FUNCTION_BLOCK FB_stringBuilder
VAR_INPUT
END_VAR
VAR
	bBuffer				:	ARRAY[0..PARAMETERS.uiMaxCharacters - 1] OF BYTE;
	bBufferOld			:	ARRAY[0..PARAMETERS.uiMaxCharacters - 1] OF BYTE;
	udiIndex			:	UDINT;
	udiIndexOld			:	UDINT;
	pbBuffer			:	POINTER TO BYTE		:=	ADR(bBuffer);
	pbBufferOld			:	POINTER TO BYTE		:=	ADR(bBufferOld);
END_VAR

METHOD AddChar : BOOL
VAR_INPUT
	byChar	:	BYTE;
END_VAR
IF CheckLength() THEN
	bBuffer[udiIndex]	:=	byChar;
	AddChar			:=	TRUE;
	IncrementIndex();
END_IF
END_METHOD

ACTION AddCloseBracket:
AddChar(41);
END_ACTION

ACTION AddColon:
AddChar(58);
END_ACTION

ACTION AddComma:
AddChar(44);
END_ACTION

ACTION AddDollar:
AddChar(36);
END_ACTION

ACTION AddDot:
AddChar(46);
END_ACTION

ACTION AddDoubleQuote:
AddChar(34);
END_ACTION

METHOD AddKeyValue : BOOL
VAR_INPUT
	psKey	:	POINTER TO STRING;
	psValue	:	POINTER TO STRING;
END_VAR
AddString(psKey);
AddColon();
AddString(psValue);
AddComma();
END_METHOD

ACTION AddNewLine:
AddChar(10);
END_ACTION

ACTION AddNullChar:
IF NOT CheckLength() THEN
	udiIndex	:=	PARAMETERS.uiMaxCharacters - 1;
END_IF
AddChar(0);
END_ACTION

ACTION AddOpenBracket:
AddChar(40);
END_ACTION

ACTION AddQuote:
AddChar(39);
END_ACTION

ACTION AddSemicolon:
AddChar(59);
END_ACTION

ACTION AddSpace:
AddChar(32);
END_ACTION

METHOD AddString : BOOL
VAR_INPUT
	psString		:	POINTER TO STRING;
END_VAR
VAR
	udiLen	:	UDINT;
END_VAR
udiLen	:=	(LEN2(psString));
IF CheckFinalLength(udiLen) THEN
	MEMCPY(pbBuffer + udiIndex, psString, udiLen);
	IncrementIndexVariable(udiLen);
	AddString	:=	TRUE;
END_IF
END_METHOD

ACTION AddTab:
AddChar(9);
END_ACTION

ACTION AddUnderscore:
AddChar(95);
END_ACTION

METHOD BuildString : BOOL
VAR_INPUT
	psString	:	POINTER TO STRING;
END_VAR
AddNullChar();
MEMCPY( psString, ADR(bBuffer), udiIndex );
END_METHOD

METHOD CheckFinalLength : BOOL
VAR_INPUT
	udiLen	:	UDINT;
END_VAR
CheckFinalLength	:=	(udiIndex + udiLen) < PARAMETERS.uiMaxCharacters;
END_METHOD

METHOD CheckLength : BOOL
VAR_INPUT
END_VAR
CheckLength	:=	CheckFinalLength(0);
END_METHOD

METHOD CheckMinimumLength : BOOL
VAR_INPUT
END_VAR
CheckMinimumLength	:=	udiIndex > 0;
END_METHOD

ACTION DecrementIndex:
IF CheckMinimumLength() THEN
	udiIndex	:=	udiIndex - 1;
END_IF
END_ACTION

METHOD DeleteChars : BOOL
VAR_INPUT
	udiNumChars	:	UDINT;
END_VAR
udiNumChars	:=	MIN(udiNumChars, udiIndex);
MEMSET(pbBuffer + (udiIndex - udiNumChars), 0, udiNumChars);
udiIndex := udiIndex - udiNumChars;
END_METHOD

ACTION IncrementIndex:
IncrementIndexVariable(1);
END_ACTION

METHOD IncrementIndexVariable : BOOL
VAR_INPUT
	udiIncrement	:	UDINT;
END_VAR
udiIndex	:=	udiIndex + udiIncrement;
END_METHOD

ACTION ResetBuffer:
IF CheckMinimumLength() THEN
	udiIndexOld	:=	udiIndex - 1;
	MEMSET(	ADR(bBufferOld), 0, PARAMETERS.uiMaxCharacters);
	MEMCPY( ADR(bBufferOld), ADR(bBuffer), udiIndexOld);
	
	ResetIndex();
	MEMSET(	ADR(bBuffer), 0, PARAMETERS.uiMaxCharacters);
END_IF
END_ACTION

ACTION ResetIndex:
udiIndex	:=	0;
END_ACTION

END_FUNCTION_BLOCK

(* stored: Version 1.1.0.1, ProductVersion 3.1.4024.9
   POU FB_stringBuilder: Id {26bce644-87e4-4374-b58f-9389bc582a26}, SpecialFunc None
   Folder ACTIONs: Id {99776992-d8a0-4ed4-aa61-350cfed19f86}
   Folder METHODs: Id {9a2113b2-3380-4328-be6b-be03ed0cc5a6}
   Method AddChar: Id {acb1b8e0-0207-4f46-8378-b68a295cf363}
   Action AddCloseBracket: Id {444bcdd4-ba94-4df4-ab4d-d2ec81607a8f}
   Action AddColon: Id {955d0969-09fd-4ef7-a5fc-925f1bf3fba6}
   Action AddComma: Id {f598045d-14ce-4e49-8860-6889173f446b}
   Action AddDollar: Id {62dc17c3-04a8-45e3-b384-0493539ef6bb}
   Action AddDot: Id {e44675ea-41f7-4475-a1a8-be67ad3f2ca2}
   Action AddDoubleQuote: Id {634a5359-7116-406e-b4c1-826d6bf2f6c9}
   Method AddKeyValue: Id {ea0220f5-ed5d-41e8-9b72-147e94feed33}
   Action AddNewLine: Id {c2c363a3-f640-4a66-9c2e-ae6cfdf7030a}
   Action AddNullChar: Id {41965dbb-6995-4e5e-9350-33895695746a}
   Action AddOpenBracket: Id {2ec56027-8c0a-434b-a7a8-c83c4f1f8e42}
   Action AddQuote: Id {a0d24b89-7c31-4ef3-9361-6e66114a55e2}
   Action AddSemicolon: Id {6e821915-2f2b-48e5-a2be-50c5a41a7f62}
   Action AddSpace: Id {efb50eb6-39f2-45ad-afb8-a2137592de0e}
   Method AddString: Id {595b4d96-b597-449d-9435-3e7e82a579a8}
   Action AddTab: Id {ee6a5a98-72fa-4ae6-9474-04a98b339a88}
   Action AddUnderscore: Id {f615e6a0-0dc8-4c8e-8542-2fb8926efc44}
   Method BuildString: Id {ca77eff2-213f-461b-8f4b-842771dfc69c}
   Method CheckFinalLength: Id {5bfcfec1-41c0-4b4b-9efc-cdfedbb5d1d9}
   Method CheckLength: Id {c6856b6b-f1b0-4936-a873-24f2736990c8}
   Method CheckMinimumLength: Id {a3deb16d-1c84-436e-9e26-91d82feaafb3}
   Action DecrementIndex: Id {80622eaf-5301-41c9-a0ec-d5673140fae2}
   Method DeleteChars: Id {9567052d-08aa-4840-a672-7ff69cd94b0e}
   Action IncrementIndex: Id {1e105e41-e1b3-4291-b4f5-b3ad8bc1f44d}
   Method IncrementIndexVariable: Id {7f43a176-ec9b-446d-98cd-00989f7ef420}
   Action ResetBuffer: Id {6fd5ed2a-147e-4efd-a713-8e4977d508a1}
   Action ResetIndex: Id {0267ccdd-742e-4881-b501-77d47e764385} *)
